(* IEC 61131-3 sources: llm-plc-st-eval/data/processed_definitivo/gemini-3.1-pro-preview/I2/zero_shot, 3 files *)

(* ---- ejec_1.st ---- *)
FUNCTION_BLOCK FB_Llenado
VAR_INPUT
    btnInicio : BOOL;
    btnParo : BOOL;
    nivelAlto : BOOL;
    nivelBajo : BOOL;
END_VAR

VAR_OUTPUT
    vLlenado : BOOL;
    motorMezcla : BOOL;
    vDescarga : BOOL;
END_VAR

VAR
    estado : INT := 0; // 0: Reposo, 1: Llenado, 2: Mezcla, 3: Descarga
    tonMezcla : TON;   // Temporizador para el motor de mezcla
END_VAR

// Lógica de paro prioritario: detiene el proceso y regresa a reposo
IF btnParo THEN
    estado := 0;
END_IF;

// Instancia del temporizador: se activa solo en el estado 2 (Mezcla)
tonMezcla(IN := (estado = 2), PT := T#60S);

// Máquina de estados del proceso
CASE estado OF
    0: // Reposo: Salidas en estado seguro (desactivadas)
        vLlenado := FALSE;
        motorMezcla := FALSE;
        vDescarga := FALSE;

        IF btnInicio THEN
            estado := 1;
        END_IF;

    1: // Llenado: Abre válvula hasta detectar nivel alto
        vLlenado := TRUE;
        motorMezcla := FALSE;
        vDescarga := FALSE;

        IF nivelAlto THEN
            estado := 2;
        END_IF;

    2: // Mezcla: Enciende motor durante 60 segundos
        vLlenado := FALSE;
        motorMezcla := TRUE;
        vDescarga := FALSE;

        IF tonMezcla.Q THEN
            estado := 3;
        END_IF;

    3: // Descarga: Abre válvula hasta detectar nivel bajo
        vLlenado := FALSE;
        motorMezcla := FALSE;
        vDescarga := TRUE;

        IF nivelBajo THEN
            estado := 0;
        END_IF;

ELSE
    // Protección contra estados inválidos
    estado := 0;
END_CASE;

END_FUNCTION_BLOCK

(* ---- ejec_2.st ---- *)
FUNCTION_BLOCK FB_Llenado
VAR_INPUT
    btnInicio : BOOL;   // Botón para iniciar el proceso
    btnParo : BOOL;     // Botón para detener el proceso y llevar a estado seguro
    nivelAlto : BOOL;   // Sensor de nivel alto
    nivelBajo : BOOL;   // Sensor de nivel bajo
END_VAR

VAR_OUTPUT
    vLlenado : BOOL;    // Válvula de llenado
    motorMezcla : BOOL; // Motor del mezclador
    vDescarga : BOOL;   // Válvula de descarga
END_VAR

VAR
    estado : INT := 0;  // Máquina de estados (0:Reposo, 1:Llenado, 2:Mezcla, 3:Descarga)
    timerMezcla : TON;  // Temporizador para la etapa de mezcla
END_VAR

// 1. Condición de paro prioritario
IF btnParo THEN
    estado := 0;
END_IF;

// 2. Máquina de estados secuencial
CASE estado OF
    0: // Etapa 0: Reposo
        IF btnInicio AND NOT btnParo THEN
            estado := 1;
        END_IF;

    1: // Etapa 1: Llenado
        IF nivelAlto THEN
            estado := 2;
        END_IF;

    2: // Etapa 2: Mezcla
        IF timerMezcla.Q THEN
            estado := 3;
        END_IF;

    3: // Etapa 3: Descarga
        IF nivelBajo THEN
            estado := 0;
        END_IF;
ELSE
    // Protección contra estados inválidos
    estado := 0;
END_CASE;

// 3. Control de salidas (Garantiza estado seguro si no es su etapa activa)
vLlenado := (estado = 1);
motorMezcla := (estado = 2);
vDescarga := (estado = 3);

// 4. Actualización del temporizador (Se activa únicamente en la etapa 2)
timerMezcla(IN := (estado = 2), PT := T#60S);

END_FUNCTION_BLOCK

(* ---- ejec_3.st ---- *)
FUNCTION_BLOCK FB_Llenado
VAR_INPUT
    btnInicio : BOOL;
    btnParo : BOOL;
    nivelAlto : BOOL;
    nivelBajo : BOOL;
END_VAR

VAR_OUTPUT
    vLlenado : BOOL;
    motorMezcla : BOOL;
    vDescarga : BOOL;
END_VAR

VAR
    estado : INT := 0; // 0: Reposo, 1: Llenado, 2: Mezcla, 3: Descarga
    tonMezcla : TON;   // Temporizador para el motor de mezcla
END_VAR

// Lógica de transición de estados y paro
IF btnParo THEN
    estado := 0; // El paro fuerza el estado de reposo
ELSE
    CASE estado OF
        0: // Etapa de Reposo
            IF btnInicio THEN
                estado := 1;
            END_IF;

        1: // Etapa de Llenado
            IF nivelAlto THEN
                estado := 2;
            END_IF;

        2: // Etapa de Mezcla
            IF tonMezcla.Q THEN
                estado := 3;
            END_IF;

        3: // Etapa de Descarga
            IF nivelBajo THEN
                estado := 0;
            END_IF;
    END_CASE;
END_IF;

// Control del temporizador (se activa solo en el estado 2)
tonMezcla(IN := (estado = 2), PT := T#60S);

// Control de salidas (al estar en estado 0 por btnParo, todas son FALSE)
vLlenado := (estado = 1);
motorMezcla := (estado = 2);
vDescarga := (estado = 3);

END_FUNCTION_BLOCK
